{attribute 'qualified_only'}
{attribute 'strict'}
TYPE E_SetJobState :
(
	eIdle := 0,
	eAxesNotReady,
	eSelNewStone,
	eSelRemoveStone,
	eCheckAllMagazines,
	eValidateNewStone,
	eValidateRemoveStone
);
END_TYPE

(* stored: Version 1.1.0.1, ProductVersion 3.1.4024.12
   DUT E_SetJobState: Id {15be2a58-62da-4ff0-b819-d961589d3a57} *)
